(* CODESYS project Glob_Var.gvl.xml

Project tree, tasks and I/O mapping:
  global variables Glob_Var
*)

// Glob_Var
{attribute 'qualified_only'}
VAR_GLOBAL
//Inputs
	TempActual: REAL:=8.0;
	TempSet: REAL:=8.0;
	DoorOpen: BOOL;
	AlarmThreshold:TIME:=T#10S;
	DoorOpenThreshold:TIME:=T#10S;

//Outputs
	Compressor: BOOL;
	Signal: BOOL;
	Lamp: BOOL;
END_VAR
